(* IEC 61131-3 sources: llm-plc-st-eval/codesys/dobles/A2, 9 files *)

(* ---- 01_Correcta.st ---- *)
(* DOBLE DE PRUEBA A2/Correcta - NO ES CORPUS. Esperado: veredicto 1 *)
FUNCTION_BLOCK FB_Batch
VAR_INPUT
    nivelA : BOOL;
    nivelB : BOOL;
    nivelVacio : BOOL;
    btnInicio : BOOL;
    btnAbort : BOOL;
    temp : REAL;
END_VAR
VAR_OUTPUT
    vA : BOOL;
    vB : BOOL;
    calentador : BOOL;
    mezclador : BOOL;
    vDescarga : BOOL;
    fase : INT;
END_VAR
VAR
    tMez : TON;
    calLat : BOOL;
END_VAR
IF btnInicio AND fase = 0 THEN
    fase := 1;
ELSIF btnAbort AND fase >= 1 AND fase <= 4 THEN
    IF nivelVacio THEN
        fase := 0;
    ELSE
        fase := 5;
    END_IF
ELSE
    CASE fase OF
        1: IF nivelA THEN fase := 2; END_IF
        2: IF nivelB THEN fase := 3; END_IF
        3: IF temp >= 60.0 THEN fase := 4; END_IF
        4: IF tMez.Q THEN fase := 5; END_IF
        5: IF nivelVacio THEN fase := 0; END_IF
    END_CASE
END_IF
tMez(IN := fase = 4, PT := T#120S);
vA := fase = 1;
vB := fase = 2;
calentador := fase = 3;
mezclador := fase = 4;
vDescarga := fase = 5;
END_FUNCTION_BLOCK

(* ---- 02_AbortEnReposo.st ---- *)
(* DOBLE DE PRUEBA A2/AbortEnReposo - NO ES CORPUS. Esperado: veredicto 2, falla en el paso 1 *)
FUNCTION_BLOCK FB_Batch
VAR_INPUT
    nivelA : BOOL;
    nivelB : BOOL;
    nivelVacio : BOOL;
    btnInicio : BOOL;
    btnAbort : BOOL;
    temp : REAL;
END_VAR
VAR_OUTPUT
    vA : BOOL;
    vB : BOOL;
    calentador : BOOL;
    mezclador : BOOL;
    vDescarga : BOOL;
    fase : INT;
END_VAR
VAR
    tMez : TON;
    calLat : BOOL;
END_VAR
IF btnAbort AND fase = 0 AND NOT nivelVacio THEN
    fase := 5;
ELSIF btnInicio AND fase = 0 THEN
    fase := 1;
ELSIF btnAbort AND fase >= 1 AND fase <= 4 THEN
    IF nivelVacio THEN
        fase := 0;
    ELSE
        fase := 5;
    END_IF
ELSE
    CASE fase OF
        1: IF nivelA THEN fase := 2; END_IF
        2: IF nivelB THEN fase := 3; END_IF
        3: IF temp >= 60.0 THEN fase := 4; END_IF
        4: IF tMez.Q THEN fase := 5; END_IF
        5: IF nivelVacio THEN fase := 0; END_IF
    END_CASE
END_IF
tMez(IN := fase = 4, PT := T#120S);
vA := fase = 1;
vB := fase = 2;
calentador := fase = 3;
mezclador := fase = 4;
vDescarga := fase = 5;
END_FUNCTION_BLOCK

(* ---- 03_InicioNoIgnorado.st ---- *)
(* DOBLE DE PRUEBA A2/InicioNoIgnorado - NO ES CORPUS. Esperado: veredicto 2, falla en el paso 5 *)
FUNCTION_BLOCK FB_Batch
VAR_INPUT
    nivelA : BOOL;
    nivelB : BOOL;
    nivelVacio : BOOL;
    btnInicio : BOOL;
    btnAbort : BOOL;
    temp : REAL;
END_VAR
VAR_OUTPUT
    vA : BOOL;
    vB : BOOL;
    calentador : BOOL;
    mezclador : BOOL;
    vDescarga : BOOL;
    fase : INT;
END_VAR
VAR
    tMez : TON;
    calLat : BOOL;
END_VAR
IF btnInicio THEN
    fase := 1;
ELSIF btnAbort AND fase >= 1 AND fase <= 4 THEN
    IF nivelVacio THEN
        fase := 0;
    ELSE
        fase := 5;
    END_IF
ELSE
    CASE fase OF
        1: IF nivelA THEN fase := 2; END_IF
        2: IF nivelB THEN fase := 3; END_IF
        3: IF temp >= 60.0 THEN fase := 4; END_IF
        4: IF tMez.Q THEN fase := 5; END_IF
        5: IF nivelVacio THEN fase := 0; END_IF
    END_CASE
END_IF
tMez(IN := fase = 4, PT := T#120S);
vA := fase = 1;
vB := fase = 2;
calentador := fase = 3;
mezclador := fase = 4;
vDescarga := fase = 5;
END_FUNCTION_BLOCK

(* ---- 04_UmbralEstricto.st ---- *)
(* DOBLE DE PRUEBA A2/UmbralEstricto - NO ES CORPUS. Esperado: veredicto 2, falla en el paso 8 *)
FUNCTION_BLOCK FB_Batch
VAR_INPUT
    nivelA : BOOL;
    nivelB : BOOL;
    nivelVacio : BOOL;
    btnInicio : BOOL;
    btnAbort : BOOL;
    temp : REAL;
END_VAR
VAR_OUTPUT
    vA : BOOL;
    vB : BOOL;
    calentador : BOOL;
    mezclador : BOOL;
    vDescarga : BOOL;
    fase : INT;
END_VAR
VAR
    tMez : TON;
    calLat : BOOL;
END_VAR
IF btnInicio AND fase = 0 THEN
    fase := 1;
ELSIF btnAbort AND fase >= 1 AND fase <= 4 THEN
    IF nivelVacio THEN
        fase := 0;
    ELSE
        fase := 5;
    END_IF
ELSE
    CASE fase OF
        1: IF nivelA THEN fase := 2; END_IF
        2: IF nivelB THEN fase := 3; END_IF
        3: IF temp > 60.0 THEN fase := 4; END_IF
        4: IF tMez.Q THEN fase := 5; END_IF
        5: IF nivelVacio THEN fase := 0; END_IF
    END_CASE
END_IF
tMez(IN := fase = 4, PT := T#120S);
vA := fase = 1;
vB := fase = 2;
calentador := fase = 3;
mezclador := fase = 4;
vDescarga := fase = 5;
END_FUNCTION_BLOCK

(* ---- 05_MezclaCorta.st ---- *)
(* DOBLE DE PRUEBA A2/MezclaCorta - NO ES CORPUS. Esperado: veredicto 2, falla en el paso 9 *)
FUNCTION_BLOCK FB_Batch
VAR_INPUT
    nivelA : BOOL;
    nivelB : BOOL;
    nivelVacio : BOOL;
    btnInicio : BOOL;
    btnAbort : BOOL;
    temp : REAL;
END_VAR
VAR_OUTPUT
    vA : BOOL;
    vB : BOOL;
    calentador : BOOL;
    mezclador : BOOL;
    vDescarga : BOOL;
    fase : INT;
END_VAR
VAR
    tMez : TON;
    calLat : BOOL;
END_VAR
IF btnInicio AND fase = 0 THEN
    fase := 1;
ELSIF btnAbort AND fase >= 1 AND fase <= 4 THEN
    IF nivelVacio THEN
        fase := 0;
    ELSE
        fase := 5;
    END_IF
ELSE
    CASE fase OF
        1: IF nivelA THEN fase := 2; END_IF
        2: IF nivelB THEN fase := 3; END_IF
        3: IF temp >= 60.0 THEN fase := 4; END_IF
        4: IF tMez.Q THEN fase := 5; END_IF
        5: IF nivelVacio THEN fase := 0; END_IF
    END_CASE
END_IF
tMez(IN := fase = 4, PT := T#60S);
vA := fase = 1;
vB := fase = 2;
calentador := fase = 3;
mezclador := fase = 4;
vDescarga := fase = 5;
END_FUNCTION_BLOCK

(* ---- 06_MezclaLarga.st ---- *)
(* DOBLE DE PRUEBA A2/MezclaLarga - NO ES CORPUS. Esperado: veredicto 2, falla en el paso 10 *)
FUNCTION_BLOCK FB_Batch
VAR_INPUT
    nivelA : BOOL;
    nivelB : BOOL;
    nivelVacio : BOOL;
    btnInicio : BOOL;
    btnAbort : BOOL;
    temp : REAL;
END_VAR
VAR_OUTPUT
    vA : BOOL;
    vB : BOOL;
    calentador : BOOL;
    mezclador : BOOL;
    vDescarga : BOOL;
    fase : INT;
END_VAR
VAR
    tMez : TON;
    calLat : BOOL;
END_VAR
IF btnInicio AND fase = 0 THEN
    fase := 1;
ELSIF btnAbort AND fase >= 1 AND fase <= 4 THEN
    IF nivelVacio THEN
        fase := 0;
    ELSE
        fase := 5;
    END_IF
ELSE
    CASE fase OF
        1: IF nivelA THEN fase := 2; END_IF
        2: IF nivelB THEN fase := 3; END_IF
        3: IF temp >= 60.0 THEN fase := 4; END_IF
        4: IF tMez.Q THEN fase := 5; END_IF
        5: IF nivelVacio THEN fase := 0; END_IF
    END_CASE
END_IF
tMez(IN := fase = 4, PT := T#180S);
vA := fase = 1;
vB := fase = 2;
calentador := fase = 3;
mezclador := fase = 4;
vDescarga := fase = 5;
END_FUNCTION_BLOCK

(* ---- 07_AbortSiempreReposo.st ---- *)
(* DOBLE DE PRUEBA A2/AbortSiempreReposo - NO ES CORPUS. Esperado: veredicto 2, falla en el paso 13 *)
FUNCTION_BLOCK FB_Batch
VAR_INPUT
    nivelA : BOOL;
    nivelB : BOOL;
    nivelVacio : BOOL;
    btnInicio : BOOL;
    btnAbort : BOOL;
    temp : REAL;
END_VAR
VAR_OUTPUT
    vA : BOOL;
    vB : BOOL;
    calentador : BOOL;
    mezclador : BOOL;
    vDescarga : BOOL;
    fase : INT;
END_VAR
VAR
    tMez : TON;
    calLat : BOOL;
END_VAR
IF btnInicio AND fase = 0 THEN
    fase := 1;
ELSIF btnAbort AND fase >= 1 AND fase <= 4 THEN
    fase := 0;
ELSE
    CASE fase OF
        1: IF nivelA THEN fase := 2; END_IF
        2: IF nivelB THEN fase := 3; END_IF
        3: IF temp >= 60.0 THEN fase := 4; END_IF
        4: IF tMez.Q THEN fase := 5; END_IF
        5: IF nivelVacio THEN fase := 0; END_IF
    END_CASE
END_IF
tMez(IN := fase = 4, PT := T#120S);
vA := fase = 1;
vB := fase = 2;
calentador := fase = 3;
mezclador := fase = 4;
vDescarga := fase = 5;
END_FUNCTION_BLOCK

(* ---- 08_AbortNoCierraCalentador.st ---- *)
(* DOBLE DE PRUEBA A2/AbortNoCierraCalentador - NO ES CORPUS. Esperado: veredicto 2, falla en el paso 21 *)
FUNCTION_BLOCK FB_Batch
VAR_INPUT
    nivelA : BOOL;
    nivelB : BOOL;
    nivelVacio : BOOL;
    btnInicio : BOOL;
    btnAbort : BOOL;
    temp : REAL;
END_VAR
VAR_OUTPUT
    vA : BOOL;
    vB : BOOL;
    calentador : BOOL;
    mezclador : BOOL;
    vDescarga : BOOL;
    fase : INT;
END_VAR
VAR
    tMez : TON;
    calLat : BOOL;
END_VAR
IF btnInicio AND fase = 0 THEN
    fase := 1;
ELSIF btnAbort AND fase >= 1 AND fase <= 4 THEN
    IF fase = 3 THEN
        calLat := TRUE;
    END_IF
    IF nivelVacio THEN
        fase := 0;
    ELSE
        fase := 5;
    END_IF
ELSE
    CASE fase OF
        1: IF nivelA THEN fase := 2; END_IF
        2: IF nivelB THEN fase := 3; END_IF
        3: IF temp >= 60.0 THEN fase := 4; END_IF
        4: IF tMez.Q THEN fase := 5; END_IF
        5: IF nivelVacio THEN fase := 0; END_IF
    END_CASE
END_IF
tMez(IN := fase = 4, PT := T#120S);
vA := fase = 1;
vB := fase = 2;
calentador := fase = 3;
mezclador := fase = 4;
vDescarga := fase = 5;
IF fase = 0 THEN
    calLat := FALSE;
END_IF
calentador := calentador OR calLat;
END_FUNCTION_BLOCK

(* ---- 09_AbortEnDescargaDetiene.st ---- *)
(* DOBLE DE PRUEBA A2/AbortEnDescargaDetiene - NO ES CORPUS. Esperado: veredicto 2, falla en el paso 13 *)
FUNCTION_BLOCK FB_Batch
VAR_INPUT
    nivelA : BOOL;
    nivelB : BOOL;
    nivelVacio : BOOL;
    btnInicio : BOOL;
    btnAbort : BOOL;
    temp : REAL;
END_VAR
VAR_OUTPUT
    vA : BOOL;
    vB : BOOL;
    calentador : BOOL;
    mezclador : BOOL;
    vDescarga : BOOL;
    fase : INT;
END_VAR
VAR
    tMez : TON;
    calLat : BOOL;
END_VAR
IF btnAbort AND fase = 5 THEN
    fase := 0;
ELSIF btnInicio AND fase = 0 THEN
    fase := 1;
ELSIF btnAbort AND fase >= 1 AND fase <= 4 THEN
    IF nivelVacio THEN
        fase := 0;
    ELSE
        fase := 5;
    END_IF
ELSE
    CASE fase OF
        1: IF nivelA THEN fase := 2; END_IF
        2: IF nivelB THEN fase := 3; END_IF
        3: IF temp >= 60.0 THEN fase := 4; END_IF
        4: IF tMez.Q THEN fase := 5; END_IF
        5: IF nivelVacio THEN fase := 0; END_IF
    END_CASE
END_IF
tMez(IN := fase = 4, PT := T#120S);
vA := fase = 1;
vB := fase = 2;
calentador := fase = 3;
mezclador := fase = 4;
vDescarga := fase = 5;
END_FUNCTION_BLOCK
